(* IEC 61131-3 sources: volt/packages/volt-lsp-iec/test-corpus/lenze-mid/Device/Plc Logic/Application/A71_LocalSources/CamControls/Pulse, 2 files *)

(* ---- fc_CamC_CP_Base.pou ---- *)
FUNCTION fc_CamC_CP_Base : BOOL
VAR_INPUT
	iEN					: BOOL;
	iStartCam			: INT;
	iMachinePosition 	: INT;
	iResetFlag			: BOOL;
END_VAR
VAR_OUTPUT

END_VAR
VAR
	tBool: BOOL;

END_VAR
VAR_IN_OUT
	ioAuxOneShot: BOOL;
END_VAR

%LANGUAGE LD
%NETWORK
ASSIGN(GE(EN := RAIL(), iMachinePosition, iStartCam).OUT AND INVERT(iResetFlag) AND iEN, Q => tBool);
%NETWORK
ASSIGN(tbool AND INVERT(ioAuxOneShot), Q => fc_CamC_CP_Base);
%NETWORK
ASSIGN(tbool, Q => ioAuxOneShot);

END_FUNCTION

(* ---- fc_CamC_CP_UDT.pou ---- *)
FUNCTION fc_CamC_CP_UDT : BOOL
VAR_INPUT
	iEN						: BOOL;
	iMachinePosition		: INT;
	iResetFlag				: BOOL;

END_VAR
VAR_OUTPUT

END_VAR
VAR

END_VAR
VAR_IN_OUT
	ioPulse	: UDT_CamPulse;
END_VAR

%LANGUAGE LD
%NETWORK
MOVE(EN := RAIL(), iMachinePosition, OUT => ioPulse.MachinePos_HMI);
%NETWORK
ASSIGN(fc_CamC_CP_Base(iEN := iEN, iStartCam := ioPulse.Start, iMachinePosition := iMachinePosition, iResetFlag := iResetFlag, ioAuxOneShot := ioPulse.OSP), Q => fc_CamC_CP_UDT, Q => ioPulse.Active);

END_FUNCTION
